(* IEC 61131-3 sources: sis-interlock-demo/tests/POUs/TruthTables/FB_VoteTableEval_Test, 12 files *)

(* ---- Eval1oo1DAMatchesModel.method.decl.st ---- *)
// AUTO-GENERATED by tools_project/gen_voting_tests.py — не редактировать: правьте генератор или модель
//   tools_project/vote_model.py и запустите python tools_project/gen_voting_tests.py
// F_VoteEval, схема 1oo1, политика DA: все 4 сочетаний состояний 1 каналов
// (требование × достоверность × запрос байпаса по каналу — для FB_Voting); ожидаемые значения —
// эталонная модель tools_project/vote_model.py. Один AssertEquals_BYTE на строку.
METHOD PRIVATE Eval1oo1DAMatchesModel
VAR
    fbRig : FB_VoteTableRig;   // стенд таблиц (новый экземпляр на тест)
    bRes  : BYTE;              // код результата строки
END_VAR

(* ---- Eval1oo1DSMatchesModel.method.decl.st ---- *)
// AUTO-GENERATED by tools_project/gen_voting_tests.py — не редактировать: правьте генератор или модель
//   tools_project/vote_model.py и запустите python tools_project/gen_voting_tests.py
// F_VoteEval, схема 1oo1, политика DS: все 4 сочетаний состояний 1 каналов
// (требование × достоверность × запрос байпаса по каналу — для FB_Voting); ожидаемые значения —
// эталонная модель tools_project/vote_model.py. Один AssertEquals_BYTE на строку.
METHOD PRIVATE Eval1oo1DSMatchesModel
VAR
    fbRig : FB_VoteTableRig;   // стенд таблиц (новый экземпляр на тест)
    bRes  : BYTE;              // код результата строки
END_VAR

(* ---- Eval1oo1VTMatchesModel.method.decl.st ---- *)
// AUTO-GENERATED by tools_project/gen_voting_tests.py — не редактировать: правьте генератор или модель
//   tools_project/vote_model.py и запустите python tools_project/gen_voting_tests.py
// F_VoteEval, схема 1oo1, политика VT: все 4 сочетаний состояний 1 каналов
// (требование × достоверность × запрос байпаса по каналу — для FB_Voting); ожидаемые значения —
// эталонная модель tools_project/vote_model.py. Один AssertEquals_BYTE на строку.
METHOD PRIVATE Eval1oo1VTMatchesModel
VAR
    fbRig : FB_VoteTableRig;   // стенд таблиц (новый экземпляр на тест)
    bRes  : BYTE;              // код результата строки
END_VAR

(* ---- Eval1oo2DAMatchesModel.method.decl.st ---- *)
// AUTO-GENERATED by tools_project/gen_voting_tests.py — не редактировать: правьте генератор или модель
//   tools_project/vote_model.py и запустите python tools_project/gen_voting_tests.py
// F_VoteEval, схема 1oo2, политика DA: все 16 сочетаний состояний 2 каналов
// (требование × достоверность × запрос байпаса по каналу — для FB_Voting); ожидаемые значения —
// эталонная модель tools_project/vote_model.py. Один AssertEquals_BYTE на строку.
METHOD PRIVATE Eval1oo2DAMatchesModel
VAR
    fbRig : FB_VoteTableRig;   // стенд таблиц (новый экземпляр на тест)
    bRes  : BYTE;              // код результата строки
END_VAR

(* ---- Eval1oo2DSMatchesModel.method.decl.st ---- *)
// AUTO-GENERATED by tools_project/gen_voting_tests.py — не редактировать: правьте генератор или модель
//   tools_project/vote_model.py и запустите python tools_project/gen_voting_tests.py
// F_VoteEval, схема 1oo2, политика DS: все 16 сочетаний состояний 2 каналов
// (требование × достоверность × запрос байпаса по каналу — для FB_Voting); ожидаемые значения —
// эталонная модель tools_project/vote_model.py. Один AssertEquals_BYTE на строку.
METHOD PRIVATE Eval1oo2DSMatchesModel
VAR
    fbRig : FB_VoteTableRig;   // стенд таблиц (новый экземпляр на тест)
    bRes  : BYTE;              // код результата строки
END_VAR

(* ---- Eval1oo2VTMatchesModel.method.decl.st ---- *)
// AUTO-GENERATED by tools_project/gen_voting_tests.py — не редактировать: правьте генератор или модель
//   tools_project/vote_model.py и запустите python tools_project/gen_voting_tests.py
// F_VoteEval, схема 1oo2, политика VT: все 16 сочетаний состояний 2 каналов
// (требование × достоверность × запрос байпаса по каналу — для FB_Voting); ожидаемые значения —
// эталонная модель tools_project/vote_model.py. Один AssertEquals_BYTE на строку.
METHOD PRIVATE Eval1oo2VTMatchesModel
VAR
    fbRig : FB_VoteTableRig;   // стенд таблиц (новый экземпляр на тест)
    bRes  : BYTE;              // код результата строки
END_VAR

(* ---- Eval2oo2DAMatchesModel.method.decl.st ---- *)
// AUTO-GENERATED by tools_project/gen_voting_tests.py — не редактировать: правьте генератор или модель
//   tools_project/vote_model.py и запустите python tools_project/gen_voting_tests.py
// F_VoteEval, схема 2oo2, политика DA: все 16 сочетаний состояний 2 каналов
// (требование × достоверность × запрос байпаса по каналу — для FB_Voting); ожидаемые значения —
// эталонная модель tools_project/vote_model.py. Один AssertEquals_BYTE на строку.
METHOD PRIVATE Eval2oo2DAMatchesModel
VAR
    fbRig : FB_VoteTableRig;   // стенд таблиц (новый экземпляр на тест)
    bRes  : BYTE;              // код результата строки
END_VAR

(* ---- Eval2oo2DSMatchesModel.method.decl.st ---- *)
// AUTO-GENERATED by tools_project/gen_voting_tests.py — не редактировать: правьте генератор или модель
//   tools_project/vote_model.py и запустите python tools_project/gen_voting_tests.py
// F_VoteEval, схема 2oo2, политика DS: все 16 сочетаний состояний 2 каналов
// (требование × достоверность × запрос байпаса по каналу — для FB_Voting); ожидаемые значения —
// эталонная модель tools_project/vote_model.py. Один AssertEquals_BYTE на строку.
METHOD PRIVATE Eval2oo2DSMatchesModel
VAR
    fbRig : FB_VoteTableRig;   // стенд таблиц (новый экземпляр на тест)
    bRes  : BYTE;              // код результата строки
END_VAR

(* ---- Eval2oo2VTMatchesModel.method.decl.st ---- *)
// AUTO-GENERATED by tools_project/gen_voting_tests.py — не редактировать: правьте генератор или модель
//   tools_project/vote_model.py и запустите python tools_project/gen_voting_tests.py
// F_VoteEval, схема 2oo2, политика VT: все 16 сочетаний состояний 2 каналов
// (требование × достоверность × запрос байпаса по каналу — для FB_Voting); ожидаемые значения —
// эталонная модель tools_project/vote_model.py. Один AssertEquals_BYTE на строку.
METHOD PRIVATE Eval2oo2VTMatchesModel
VAR
    fbRig : FB_VoteTableRig;   // стенд таблиц (новый экземпляр на тест)
    bRes  : BYTE;              // код результата строки
END_VAR

(* ---- Eval2oo3DAMatchesModel.method.decl.st ---- *)
// AUTO-GENERATED by tools_project/gen_voting_tests.py — не редактировать: правьте генератор или модель
//   tools_project/vote_model.py и запустите python tools_project/gen_voting_tests.py
// F_VoteEval, схема 2oo3, политика DA: все 64 сочетаний состояний 3 каналов
// (требование × достоверность × запрос байпаса по каналу — для FB_Voting); ожидаемые значения —
// эталонная модель tools_project/vote_model.py. Один AssertEquals_BYTE на строку.
METHOD PRIVATE Eval2oo3DAMatchesModel
VAR
    fbRig : FB_VoteTableRig;   // стенд таблиц (новый экземпляр на тест)
    bRes  : BYTE;              // код результата строки
END_VAR

(* ---- Eval2oo3DSMatchesModel.method.decl.st ---- *)
// AUTO-GENERATED by tools_project/gen_voting_tests.py — не редактировать: правьте генератор или модель
//   tools_project/vote_model.py и запустите python tools_project/gen_voting_tests.py
// F_VoteEval, схема 2oo3, политика DS: все 64 сочетаний состояний 3 каналов
// (требование × достоверность × запрос байпаса по каналу — для FB_Voting); ожидаемые значения —
// эталонная модель tools_project/vote_model.py. Один AssertEquals_BYTE на строку.
METHOD PRIVATE Eval2oo3DSMatchesModel
VAR
    fbRig : FB_VoteTableRig;   // стенд таблиц (новый экземпляр на тест)
    bRes  : BYTE;              // код результата строки
END_VAR

(* ---- Eval2oo3VTMatchesModel.method.decl.st ---- *)
// AUTO-GENERATED by tools_project/gen_voting_tests.py — не редактировать: правьте генератор или модель
//   tools_project/vote_model.py и запустите python tools_project/gen_voting_tests.py
// F_VoteEval, схема 2oo3, политика VT: все 64 сочетаний состояний 3 каналов
// (требование × достоверность × запрос байпаса по каналу — для FB_Voting); ожидаемые значения —
// эталонная модель tools_project/vote_model.py. Один AssertEquals_BYTE на строку.
METHOD PRIVATE Eval2oo3VTMatchesModel
VAR
    fbRig : FB_VoteTableRig;   // стенд таблиц (новый экземпляр на тест)
    bRes  : BYTE;              // код результата строки
END_VAR
